Fanuc KAREL source: kc00009.KL

-- PROVISIONAL review KL for V1013-1; original PC SHA256 7dc4e9466fd0686ee3abf0f163fcd80030bf4def01f41b0e445b50a55a48f158
-- Incomplete behavior may be omitted. Consult companion uncertainty JSON. Do not deploy.
PROGRAM KC00009
%NOLOCKGROUP
BEGIN
  -- UNRESOLVED_PC offsets 5-33; opcodes 27,22,1C,22,22,31
  -- UNRESOLVED_PC offsets 38-42; opcodes 7F
END KC00009
